// TIA Portal V21 export
// export: Created 2026-11-21T10:55:44.8884934Z, ExportSetting WithDefaults, DisplayName Totally Integrated Automation Portal, DisplayVersion V21, DisplayName STEP 7 Professional, DisplayVersion V21, DisplayName STEP 7 Safety, DisplayVersion V21, DisplayName Tech WebApplication, DisplayVersion V21, DisplayName WinCC Basic/Comfort/Advanced, DisplayVersion V21, DisplayName WinCC Unified, DisplayVersion V21
VAR_GLOBAL   // PLC tag table "Beschriftung"
   Lamp_Überlast AT %Q0.0 : Bool;   // Überlast der Pumpe – Leuchte
   Sensor_Niveau AT %IW2 : Int;   // Capteur de niveau, en ‰
   Etikett AT %MW4 : Word;   // ラベル番号 (標識)
END_VAR
